// TIA Portal V20 export
// export: Created 2026-10-12T16:46:22.6949063Z, ExportSetting WithDefaults, DisplayName Totally Integrated Automation Portal, DisplayVersion V20 Update 6, DisplayName TIA Portal Openness, DisplayVersion V20 Update 6, DisplayName TIA Portal Version Control Interface, DisplayVersion V20 Update 6, DisplayName SINAMICS Startdrive Advanced, DisplayVersion V20 SP1 Update 2, DisplayName SINAMICS Startdrive G110M, G120, G120C, G120D, G120P, G115D, DisplayVersion V20 SP1 Update 2, DisplayName SINAMICS Startdrive G130, G150, S120, S150, SINAMICS MV, G220, S200, S210, DisplayVersion V20 SP1 Update 2, DisplayName STEP 7 Professional, DisplayVersion V20 Update 6, DisplayName STEP 7 Safety, DisplayVersion V20 Update 2, DisplayName WinCC Basic/Comfort/Advanced, DisplayVersion V20 Update 6, DisplayName WinCC Professional, DisplayVersion V20 Update 6, DisplayName WinCC Unified, DisplayVersion V20 Update 6
TYPE "UDT_FK_IN"
// stored: IsFailsafeCompliant false
   STRUCT
      Reserved : Word;   // Byte 0-1
      Status : Word;   // Byte 2-3: StatusRegister
      Warnings : Word;   // Byte 4-5: WarningsRegister
      Alarms : Word;   // Byte 6-7: AlarmsRegsiter
      ActVoltage : Int;   // Byte 8-9: x0,01V
      ActCurrent : Int;   // Byte 10-11: x1A
      Padding : Array[0..9] of Word;   // Byte 12-31: Ungenutzt
   END_STRUCT;
END_TYPE
